KUKA KRL program: ThreadProg.src

DEF ThreadProg()
; Program generated by RoboDK v5.9.4 for R1 on 26/10/2026 01:01:11
; Using nominal kinematics.
BAS(#INITMOV,0)
$ORI_TYPE  = #VAR
$CIRC_TYPE = #BASE
$VEL.ORI1 = 200
$VEL.ORI2 = 200
$ACC.ORI1 = 100
$ACC.ORI2 = 100
$ADVANCE = 2
$ACT_EX_AX = 0
PTP $AXIS_ACT ; skip BCO quickly
$BASE = {FRAME: X 1671.225,Y -0.000,Z 1507.335,A 30.000,B 0.000,C 0.000}
$TOOL = {FRAME: X 0.000,Y 0.000,Z 120.000,A 0.000,B 15.000,C 0.000}
; Thread body
END
